(* IEC 61131-3 sources: CS_4_Aufzugsteuerung/src/Stations/CP112/Steuerung/Class/SafetyBaseFSoE (part 6) *)

END_FUNCTION

FUNCTION SafetyBaseFSoE::AddToCache
  VAR_INPUT
    p_SDORequestBuffer 	: ^SDORequReadConfig;
    p_SDOResponseBuffer 	: ^SDORespReadConfig;
  END_VAR

  if p_SDORequestBuffer^.us_Length then
    CachedAddr := p_SDORequestBuffer^.ud_Address;
    CachedSize := p_SDORequestBuffer^.us_Length;
    _memcpy(ptr1:=#Cache, ptr2:=#p_SDOResponseBuffer^.ud_Data, cntr:=p_SDORequestBuffer^.us_Length);
  end_if;

END_FUNCTION

FUNCTION SafetyBaseFSoE::GetFSoEConnectionInfos
  VAR_INPUT
    p_SDORequestBuffer 	: ^SafetyBaseFSoE::SDORequReadConfig;
    p_SDOResponseBuffer 	: ^SafetyBaseFSoE::SDORespReadConfig;
  END_VAR
  VAR
    Address         : UDINT;
    Size            : USINT;
    sd_retval       : DINT;
    i               : UDINT;
    pActConnection  : ^t_FSoEConnectionDetails;
    TempRoutingInfo : t_FSoERoutingInfoElement;
    NextAddress     : UDINT;
  END_VAR

  // always free the connection infos
  FreeFSoEConnectionInfos(bFreeAlways:=TRUE);

  // check if we already got the info:
  if ConnectionInfos.ConnectionNo | ConnectionInfos.pFirstConnection then
    LogError("@0280 (SafetyBaseFSoE::GetFSoEConnectionInfos) List already exists! May not have been resetted correctly!");
    return;
  end_if;

//*****************************************************************************
//** CONNECTION STATE INFO                                                   **
//*****************************************************************************

  // get number of connections
  Address := SBF_SDO_ADDRESS_FSOE_CONN_STATE;
  Size    := 2;

  //send request and receive data
  sd_retval := SDOReadCfgRequ ( p_SDORequestBuffer  := p_SDORequestBuffer
                              , p_SDOResponseBuffer := p_SDOResponseBuffer
                              , ud_Address          := Address
                              , us_Length           := Size
                              );

  //no response
  if ( sd_retval <> 0 ) then
    LogError("@0281 (SafetyBaseFSoE::GetFSoEConnectionInfos) Error reading number of connections.");
    return;
  end_if;

  ConnectionInfos.ConnectionNo := p_SDOResponseBuffer^.ud_Data$UINT;

  if ConnectionInfos.ConnectionNo = 0 then
    // no connections available
    return;
  end_if;

  // allocate memory for the connections
  ConnectionInfos.pFirstConnection$pVoid := ToStdLib.Malloc(size:= ConnectionInfos.ConnectionNo * sizeof(t_FSoEConnectionDetails));

  if ConnectionInfos.pFirstConnection = NIL then
    LogError("@0282 (SafetyBaseFSoE::GetFSoEConnectionInfos) Failed to allocate memory for FSoE connection details.");
    return;
  end_if;

  // reset memory (also resets pNext although we are not using a linked list here)
  _memset(dest:=ConnectionInfos.pFirstConnection, usByte:=0, cntr:= ConnectionInfos.ConnectionNo * sizeof(t_FSoEConnectionDetails));

  Address += Size;
  Size    := 1;

  pActConnection := ConnectionInfos.pFirstConnection;

  // get connection states
  for i := 0 to ConnectionInfos.ConnectionNo-1 do
    // get state of connection

    //send request and receive data
    sd_retval := SDOReadCfgRequ ( p_SDORequestBuffer  := p_SDORequestBuffer
                                , p_SDOResponseBuffer := p_SDOResponseBuffer
                                , ud_Address          := Address
                                , us_Length           := Size
                                );

    //no response
    if ( sd_retval <> 0 ) then
      LogError("@0283 (SafetyBaseFSoE::GetFSoEConnectionInfos) Error reading connection state.");
      return;
    end_if;

    // get connection state
    pActConnection^.ConnectionState := (p_SDOResponseBuffer^.ud_Data$USINT AND 2#0111)$t_FSoEConnectionState;

    // get info if the module is master or slave at this connection
    pActConnection^.Flags.IsMaster  := (p_SDOResponseBuffer^.ud_Data$USINT AND 2#1000) <> 0;

    // save safety number
    pActConnection^.OwnerSafetyNbr  := SafetyNumber;

    // for easier debugging we set the correct next pointers
    if i = ConnectionInfos.ConnectionNo-1 then
      pActConnection^.pNext := NIL;
    else
      pActConnection^.pNext := pActConnection + sizeof(t_FSoEConnectionDetails);
    end_if;

    pActConnection                  += sizeof(t_FSoEConnectionDetails);
    Address                         += Size;
  end_for;

//*****************************************************************************
//** ROUTING INFO                                                            **
//*****************************************************************************

  // get number of connections
  Address := SBF_SDO_ADDRESS_FSOE_ROUTING_INFO;
  Size    := 2;

  //send request and receive data
  sd_retval := SDOReadCfgRequ ( p_SDORequestBuffer  := p_SDORequestBuffer
                              , p_SDOResponseBuffer := p_SDOResponseBuffer
                              , ud_Address          := Address
                              , us_Length           := Size
                              );

  //no response
  if ( sd_retval <> 0 ) then
    LogError("@0281 (SafetyBaseFSoE::GetFSoEConnectionInfos) Error reading number of connections.");
    return;
  end_if;

  // check if it's the same number
  if ConnectionInfos.ConnectionNo <> p_SDOResponseBuffer^.ud_Data$UINT then
    LogError("@0285 (SafetyBaseFSoE::GetFSoEConnectionInfos) Number of connections does not match (case 1).");
    return;
  end_if;

  Address += Size;
  Size    := sizeof(t_FSoERoutingInfoElement);

  pActConnection := ConnectionInfos.pFirstConnection;

  // get connection states
  for i := 0 to ConnectionInfos.ConnectionNo-1 do
    // get routing info of connections

    //send request and receive data
    sd_retval := SDOReadCfgRequ ( p_SDORequestBuffer  := p_SDORequestBuffer
                                , p_SDOResponseBuffer := p_SDOResponseBuffer
                                , ud_Address          := Address
                                , us_Length           := Size
                                );

    //no response
    if ( sd_retval <> 0 ) then
      LogError("@0286 (SafetyBaseFSoE::GetFSoEConnectionInfos) Error reading routing info.");
      return;
    end_if;

    TempRoutingInfo := p_SDOResponseBuffer^.ud_Data$t_FSoERoutingInfoElement;

    // store the data in the connection info
    pActConnection^.SlaveAddress        := TempRoutingInfo.SlaveAddress;
    pActConnection^.MasterReadSize      := TempRoutingInfo.SafeOutputFrameSize;
    pActConnection^.MasterWriteSize     := TempRoutingInfo.SafeInputFrameSize;

    // the offset info depends on if we are master or slave
    if pActConnection^.Flags.IsMaster then
      pActConnection^.MasterReadOffset  := TempRoutingInfo.SafeOutputFrameOffset;
      pActConnection^.MasterWriteOffset := TempRoutingInfo.SafeInputFrameOffset;
    else
      pActConnection^.SlaveWriteOffset  := TempRoutingInfo.SafeOutputFrameOffset;
      pActConnection^.SlaveReadOffset   := TempRoutingInfo.SafeInputFrameOffset;
    end_if;

    pActConnection                  += sizeof(t_FSoEConnectionDetails);
    Address                         += Size;
  end_for;

//*****************************************************************************
//** CONNECTION INSTANCES                                                    **
//*****************************************************************************

  Address := SBF_SDO_ADDRESS_FSOE_CONN_INST;
  Size    := 4;

  //send request and receive data
  sd_retval := SDOReadCfgRequ ( p_SDORequestBuffer  := p_SDORequestBuffer
                              , p_SDOResponseBuffer := p_SDOResponseBuffer
                              , ud_Address          := Address
                              , us_Length           := Size
                              );

  //no response
  if ( sd_retval <> 0 ) then
    LogError("@0281 (SafetyBaseFSoE::GetFSoEConnectionInfos) Error reading number of connections.");
    return;
  end_if;

  // check if it's the same number
  if ConnectionInfos.ConnectionNo <> p_SDOResponseBuffer^.ud_Data then
    LogError("@0287 (SafetyBaseFSoE::GetFSoEConnectionInfos) Number of connections does not match (case 2).");
    return;
  end_if;

  Address += Size;

  pActConnection := ConnectionInfos.pFirstConnection;

  // get connection states
  for i := 0 to ConnectionInfos.ConnectionNo-1 do
    // get routing instance info of connections

    Size := 4;

    //send request and receive data
    sd_retval := SDOReadCfgRequ ( p_SDORequestBuffer  := p_SDORequestBuffer
                                , p_SDOResponseBuffer := p_SDOResponseBuffer
                                , ud_Address          := Address
                                , us_Length           := Size
                                );

    //no response
    if ( sd_retval <> 0 ) then
      LogError("@0288 (SafetyBaseFSoE::GetFSoEConnectionInfos) Error reading size of routing instance info.");
      return;
    end_if;

    // calculate address of next connection (to check it later)
    NextAddress := Address + p_SDOResponseBuffer^.ud_Data;

    // get the flags
    Address   += Size;
    Size      := 4;

    //send request and receive data
    sd_retval := SDOReadCfgRequ ( p_SDORequestBuffer  := p_SDORequestBuffer
                                , p_SDOResponseBuffer := p_SDOResponseBuffer
                                , ud_Address          := Address
                                , us_Length           := Size
                                );

    //no response
    if ( sd_retval <> 0 ) then
      LogError("@0289 (SafetyBaseFSoE::GetFSoEConnectionInfos) Error reading flags of routing instance info.");
      return;
    end_if;

    if ((p_SDOResponseBuffer^.ud_Data AND 1) <> 0) <> pActConnection^.Flags.IsMaster then
      LogError("@028A (SafetyBaseFSoE::GetFSoEConnectionInfos) Master settings mismatch.");
      return;
    end_if;

    //! Flags
    //  Actually, type is 4 bytes in size but for compatibility reasons it is still used as 1 byte. As a result, bits 9-32 are currently not used.
    //  Bit1: 1, wenn FSoE-Master, 0=FSoE-Slave
    //  Bit2: 1, wenn die Slave-Adresse über den HW-Pfad ermittelt wird
    //  Bit3: 1, wenn CRC von der FW ermittelt werden muss
    //  Bit4: 1, wenn Interface und Slave
    //  Bit5: 1, wenn Multichannel verwendet werden, aber ein Multichannel ist nicht vorhanden und der Eingang auf 1 gesetzt wird.
    //  Bit6: 1, wenn der Adressvergabeservice verwendet werden soll
    //  Bit7: 1, wenn der Master beim Slave die Connection ID anfordert
    //  Bit8: 1, wenn es sich um ein HGW handelt
    //  Bit9: 1, wenn Assign Slave On Demand
    //  Bits 10-32: reserviert, sind auf 0 gesetzt und werden nicht ausgewertet

    //check size of FSoEFlags type --> possible are 1 or 4 byte
    pActConnection^.Flags := p_SDOResponseBuffer^.ud_Data$t_FSoEFlags;

    if (pActConnection^.Flags AND SM_FLAGS_FLEXCON_MASK) = SM_FLAGS_FLEXCON_NODE then
#ifdef SAFETY_DEBUG_LOGGING_ACTIVATED
      LogError(e_msg:="SafetyBaseFSoE: Found FSOE Connection of FlexConNode");
#endif
      sFlexCon.FoundNodeInConfig := TRUE;
    elsif (pActConnection^.Flags AND SM_FLAGS_FLEXCON_MASK) = SM_FLAGS_FLEXCON_HOST then
#ifdef SAFETY_DEBUG_LOGGING_ACTIVATED
      LogError(e_msg:="SafetyBaseFSoE: Found FSOE Connection of FlexConHost");
#endif
      sFlexCon.FoundHostInConfig := TRUE;
    end_if;

    // get the net size of the safe output data (only the bits for the I/Os without crc and stuff)
    Address   += Size;
    Size      := 2;

    //send request and receive data
    sd_retval := SDOReadCfgRequ ( p_SDORequestBuffer  := p_SDORequestBuffer
                                , p_SDOResponseBuffer := p_SDOResponseBuffer
                                , ud_Address          := Address
                                , us_Length           := Size
                                );

    //no response
    if ( sd_retval <> 0 ) then
      LogError("@028B (SafetyBaseFSoE::GetFSoEConnectionInfos) Error reading safe output net size of routing instance info.");
      return;
    end_if;

    // we don't need the net size yet

    // get the net size of the safe input data (only the bits for the I/Os without crc and stuff)
    Address   += Size;
    Size      := 2;

    //send request and receive data
    sd_retval := SDOReadCfgRequ ( p_SDORequestBuffer  := p_SDORequestBuffer
                                , p_SDOResponseBuffer := p_SDOResponseBuffer
                                , ud_Address          := Address
                                , us_Length           := Size
                                );

    //no response
    if ( sd_retval <> 0 ) then
      LogError("@028C (SafetyBaseFSoE::GetFSoEConnectionInfos) Error reading safe input net size of routing instance info.");
      return;
    end_if;

    // we don't need the net size yet

    // get the slave address
    Address   += Size;
    Size      := 2;

    //send request and receive data
    sd_retval := SDOReadCfgRequ ( p_SDORequestBuffer  := p_SDORequestBuffer
                                , p_SDOResponseBuffer := p_SDOResponseBuffer
                                , ud_Address          := Address
                                , us_Length           := Size
                                );

    //no response
    if ( sd_retval <> 0 ) then
      LogError("@028D (SafetyBaseFSoE::GetFSoEConnectionInfos) Error reading slave address of routing instance info.");
      return;
    end_if;

    // the following settings are only available in the master
    if pActConnection^.Flags.IsMaster then

      // get the connection ID
      Address   += Size;
      Size      := 2;

      //send request and receive data
      sd_retval := SDOReadCfgRequ ( p_SDORequestBuffer  := p_SDORequestBuffer
                                  , p_SDOResponseBuffer := p_SDOResponseBuffer
                                  , ud_Address          := Address
                                  , us_Length           := Size
                                  );

      //no response
      if ( sd_retval <> 0 ) then
        LogError("@028E (SafetyBaseFSoE::GetFSoEConnectionInfos) Error reading the connection ID of routing instance info.");
        return;
      end_if;

      pActConnection^.ConnectionID := p_SDOResponseBuffer^.ud_Data$UINT;

      // get transmission time
      Address   += Size;
      Size      := 2;

      //send request and receive data
      sd_retval := SDOReadCfgRequ ( p_SDORequestBuffer  := p_SDORequestBuffer
                                  , p_SDOResponseBuffer := p_SDOResponseBuffer
                                  , ud_Address          := Address
                                  , us_Length           := Size
                                  );

      //no response
      if ( sd_retval <> 0 ) then
        LogError("@028F (SafetyBaseFSoE::GetFSoEConnectionInfos) Error reading the transmission time of routing instance info.");
        return;
      end_if;

      pActConnection^.TransmissionTime_ms := p_SDOResponseBuffer^.ud_Data$UINT;

      // get length of communication parameters (must be 2)
      Address   += Size;
      Size      := 2;

      //send request and receive data
      sd_retval := SDOReadCfgRequ ( p_SDORequestBuffer  := p_SDORequestBuffer
                                  , p_SDOResponseBuffer := p_SDOResponseBuffer
                                  , ud_Address          := Address
                                  , us_Length           := Size
                                  );

      //no response
      if ( sd_retval <> 0 ) then
        LogError("@0290 (SafetyBaseFSoE::GetFSoEConnectionInfos) Error reading the length of the communication parameters of routing instance info.");
        return;
      end_if;

      if p_SDOResponseBuffer^.ud_Data$UINT <> 2 then
        LogError("@0291 (SafetyBaseFSoE::GetFSoEConnectionInfos) Length of communication parameters is wrong.");
        return;
      end_if;

      // skip FSoE watchdog time in ms
      Address   += Size;
      Size      := 2;

      // get size of application parameters
      Address   += Size;
      Size      := 2;

      //send request and receive data
      sd_retval := SDOReadCfgRequ ( p_SDORequestBuffer  := p_SDORequestBuffer
                                  , p_SDOResponseBuffer := p_SDOResponseBuffer
                                  , ud_Address          := Address
                                  , us_Length           := Size
                                  );

      //no response
      if ( sd_retval <> 0 ) then
        LogError("@0292 (SafetyBaseFSoE::GetFSoEConnectionInfos) Error reading the length of the application parameters of routing instance info.");
        return;
      end_if;

      // skip length
      Address   += Size;

      // skip application parameters
      Size      := p_SDOResponseBuffer^.ud_Data$USINT;
      Address   += Size;

      // get to a 4 byte aligned address
      if (Address MOD 4) then
        Address := Address + (4 - (Address MOD 4)); //increase memory, up to a value, which could be divided by 4
      end_if;

      // get size of hw path
      Size      := 4;

      //send request and receive data
      sd_retval := SDOReadCfgRequ ( p_SDORequestBuffer  := p_SDORequestBuffer
                                  , p_SDOResponseBuffer := p_SDOResponseBuffer
                                  , ud_Address          := Address
                                  , us_Length           := Size
                                  );

      //no response
      if ( sd_retval <> 0 ) then
        LogError("@0293 (SafetyBaseFSoE::GetFSoEConnectionInfos) Error reading the hardware path length of routing instance info.");
        return;
      end_if;

      // get the hardware path
      Address   += Size;
      Size      := p_SDOResponseBuffer^.ud_Data$USINT;

      if Size = 0 then
        LogError("@0294 (SafetyBaseFSoE::GetFSoEConnectionInfos) Hardware path length is zero.");
        return;
      end_if;

      //send request and receive data
      sd_retval := SDOReadCfgRequ ( p_SDORequestBuffer  := p_SDORequestBuffer
                                  , p_SDOResponseBuffer := p_SDOResponseBuffer
                                  , ud_Address          := Address
                                  , us_Length           := Size
                                  );

      //no response
      if ( sd_retval <> 0 ) then
        LogError("@0295 (SafetyBaseFSoE::GetFSoEConnectionInfos) Error reading the hardware path of routing instance info.");
        return;
      end_if;

      // save hardware path into structure
      pActConnection^.SlavePathLen      := Size;
      pActConnection^.pSlavePath$pVoid  := ToStdLib.Malloc(size:=Size);

      if pActConnection^.pSlavePath = NIL then
        LogError("@0296 (SafetyBaseFSoE::GetFSoEConnectionInfos) Failed to allocate memory for the slave hardware path at the routing instance info.");
        return;
      end_if;

      _memcpy(ptr1:=pActConnection^.pSlavePath, ptr2:=#p_SDOResponseBuffer^.ud_Data, cntr:=pActConnection^.SlavePathLen);

      Address         += Size;

      // get to a 4 byte aligned address
      if (Address MOD 4) then
        Address := Address + (4 - (Address MOD 4)); //increase memory, up to a value, which could be divided by 4
      end_if;

      // get size of compressed hw path
      Size      := 4;

      //send request and receive data
      sd_retval := SDOReadCfgRequ ( p_SDORequestBuffer  := p_SDORequestBuffer
                                  , p_SDOResponseBuffer := p_SDOResponseBuffer
                                  , ud_Address          := Address
                                  , us_Length           := Size
                                  );

      //no response
      if ( sd_retval <> 0 ) then
        LogError("@0297 (SafetyBaseFSoE::GetFSoEConnectionInfos) Error reading the compressed hardware path length of routing instance info.");
        return;
      end_if;

      // get the hardware path
      Address   += Size;
      Size      := p_SDOResponseBuffer^.ud_Data$USINT;

      //send request and receive data
      sd_retval := SDOReadCfgRequ ( p_SDORequestBuffer  := p_SDORequestBuffer
                                  , p_SDOResponseBuffer := p_SDOResponseBuffer
                                  , ud_Address          := Address
                                  , us_Length           := Size
                                  );

      //no response
      if ( sd_retval <> 0 ) then
        LogError("@0298 (SafetyBaseFSoE::GetFSoEConnectionInfos) Error reading the compressed hardware path of routing instance info.");
        return;
      end_if;

      // save compressed hardware path into structure
      pActConnection^.SlavePathCompLen      := Size;
      pActConnection^.pSlavePathComp$pVoid  := ToStdLib.Malloc(size:=Size);

      if pActConnection^.pSlavePathComp = NIL then
        LogError("@0299 (SafetyBaseFSoE::GetFSoEConnectionInfos) Failed to allocate memory for the compressed slave hardware path at the routing instance info.");
        return;
      end_if;

      _memcpy(ptr1:=pActConnection^.pSlavePathComp, ptr2:=#p_SDOResponseBuffer^.ud_Data, cntr:=pActConnection^.SlavePathCompLen);

      if  (pActConnection^.pSlavePathComp^ = 6) &
          ((pActConnection^.pSlavePathComp + 5)^$HDINT AND 16#00FFFFFF) = 0 then

        // special IP: (0.0.0.x)
        // if custom ip is detected change pathcomp type from 6 (IP) to 3 (Interface)
        pActConnection^.pSlavePathComp^ :=3;
      end_if;

      //Get slot ID and communication ID from HGW
      if pActConnection^.Flags.IsHGW then

        //Get machinenumber of FUB
        sd_retval := SDOReadCfgRequ ( p_SDORequestBuffer  := p_SDORequestBuffer
                                    , p_SDOResponseBuffer := p_SDOResponseBuffer
                                    , ud_Address          := SBF_SDO_ADDRESS_HGW_FUB_BASE_ADDRESS + SBF_SDO_ADDRESS_HGW_OFFSET_MACHINENUMBER
                                    , us_Length           := 4
                                    , b_UseCache          := FALSE
                                    );

        //no response
        if ( sd_retval <> 0 ) then
          LogError("@03DA (SafetyBaseFSoE::GetFSoEConnectionInfos) Error reading the machinenumber of routing instance info.");
          return;
        end_if;

        sHGW.udMachineNrb := p_SDOResponseBuffer^.ud_Data$UDINT;

        // get the Slot ID
        Address   += Size;
        Size      := 2;

        //send request and receive data
        sd_retval := SDOReadCfgRequ ( p_SDORequestBuffer  := p_SDORequestBuffer
                                    , p_SDOResponseBuffer := p_SDOResponseBuffer
                                    , ud_Address          := Address
                                    , us_Length           := Size
                                    );

        //no response
        if ( sd_retval <> 0 ) then
          LogError("@03DB (SafetyBaseFSoE::GetFSoEConnectionInfos) Error reading the communication ID of routing instance info.");
          return;
        end_if;

        sHGW.uiCommunicationID := p_SDOResponseBuffer^.ud_Data$UINT;

        // get the communication ID
        Address   += Size;
        Size      := 2;

        //send request and receive data
        sd_retval := SDOReadCfgRequ ( p_SDORequestBuffer  := p_SDORequestBuffer
                                    , p_SDOResponseBuffer := p_SDOResponseBuffer
                                    , ud_Address          := Address
                                    , us_Length           := Size
                                    );

        //no response
        if ( sd_retval <> 0 ) then
          LogError("@03DC (SafetyBaseFSoE::GetFSoEConnectionInfos) Error reading the slot ID of routing instance info.");
          return;
        end_if;

        sHGW.uiSlotID := p_SDOResponseBuffer^.ud_Data$UINT;

        //save fsoe pdo offsets and length
        sHGW.InputPDOLength  := pActConnection^.MasterWriteSize;
        sHGW.OutputPDOLength := pActConnection^.MasterReadSize;
        if pActConnection^.Flags.IsMaster then
          sHGW.InputPDOOffset  := pActConnection^.MasterWriteOffset;
          sHGW.OutputPDOOffset := pActConnection^.MasterReadOffset;
        else
          sHGW.InputPDOOffset  := pActConnection^.SlaveWriteOffset;
          sHGW.OutputPDOOffset := pActConnection^.SlaveReadOffset;
        end_if;
        sHGW.uiTransmissionTime_ms := pActConnection^.TransmissionTime_ms;
      end_if;

      Address         += Size;

      // get to a 4 byte aligned address
      if (Address MOD 4) then
        Address := Address + (4 - (Address MOD 4)); //increase memory, up to a value, which could be divided by 4
      end_if;

      if Address > NextAddress then
        LogError("@029A (SafetyBaseFSoE::GetFSoEConnectionInfos) Structure size mismatch.");
        return;
      end_if;
    end_if;

    Address         := NextAddress;
    pActConnection  += sizeof(t_FSoEConnectionDetails);
  end_for;

END_FUNCTION

FUNCTION SafetyBaseFSoE::FreeFSoEConnectionInfos
	VAR_INPUT
		bFreeAlways 	: BOOL;(* := false *)
	END_VAR
  VAR
    i               : UDINT;
    pActConnection  : ^t_FSoEConnectionDetails;
  END_VAR

  if (ConnectionInfos.ConnectionNo = 0) | (ConnectionInfos.pFirstConnection = NIL) then
    // nothing to free
    return;
  end_if;

  //Check if we want to clear the connection infos always
  if bFreeAlways = false then
    // check if all connections have been initialized
    pActConnection := ConnectionInfos.pFirstConnection;
    for i := 0 to ConnectionInfos.ConnectionNo-1 do
      if pActConnection^.ConnectionState = FCS_NOT_INITIALIZED then
        // not yet time to free them
        return;
      end_if;

      pActConnection += sizeof(t_FSoEConnectionDetails);
    end_for;
  end_if;

  pActConnection := ConnectionInfos.pFirstConnection;
  for i := 0 to ConnectionInfos.ConnectionNo-1 do
    // free hardware path memory

    if pActConnection^.pSlavePath then
      ToStdLib.Free(mptr:=pActConnection^.pSlavePath);
    end_if;

    if pActConnection^.pSlavePathComp then
      ToStdLib.Free(mptr:=pActConnection^.pSlavePathComp);
    end_if;

    pActConnection += sizeof(t_FSoEConnectionDetails);
  end_for;

  // free the connectionlist
  ToStdLib.Free(mptr:=ConnectionInfos.pFirstConnection);
  ConnectionInfos.pFirstConnection := NIL;
  ConnectionInfos.ConnectionNo := 0;

END_FUNCTION

FUNCTION SafetyBaseFSoE::CheckFSoEConnections
  VAR
    MyPara 	            : CmdStruct;
    MyResult	          : results;
    i                   : UDINT;
    pActConnection      : ^t_FSoEConnectionDetails;
    SDORequestBuffer    : SDORequReadConfig;
    SDOResponseBuffer   : ARRAY [0..SBF_SDO_MAX_LENGTH-1] OF USINT;
    p_SDORequestBuffer 	: ^SDORequReadConfig;
    p_SDOResponseBuffer : ^SDORespReadConfig;
    UnInifializedNo     : UDINT;
    sd_retval           : DINT;
  END_VAR

  // there were some of the FSoE connections not initialized when fetching the configuration data => update them

  UnInifializedNo := 0;

  //SDO request for this command has 5 bytes additional to the header
  p_SDORequestBuffer := #SDORequestBuffer;

  //SDO response for this command can have maximum additional data
  p_SDOResponseBuffer := (#SDOResponseBuffer)$^SDORespReadConfig;

  //calculate length without crc
  p_SDORequestBuffer^.StdHeader.Len := sizeof(SDORequReadConfig) - sizeof(SDOHeader.StdHeader.CRC);

  //type
  p_SDORequestBuffer^.StdHeader.Typ := SDO_STD;

  //command for reading config data
  p_SDORequestBuffer^.StdHeader.Cmd := SBF_SDO_COMMAND_READ;

  // reset cache, because it may contain an old access on the same address => we want fresh data
  CachedSize := 0;

  pActConnection := ConnectionInfos.pFirstConnection;

  for i := 0 to ConnectionInfos.ConnectionNo-1 do
    if pActConnection^.ConnectionState = FCS_NOT_INITIALIZED then
      UnInifializedNo += 1;

      //send request and receive data
      sd_retval := SDOReadCfgRequ ( p_SDORequestBuffer  := p_SDORequestBuffer
                                  , p_SDOResponseBuffer := p_SDOResponseBuffer
                                  , ud_Address          := SBF_SDO_ADDRESS_FSOE_CONN_STATE + 2 + i
                                  , us_Length           := 1
                                  );

      //no response
      if ( sd_retval <> 0 ) then
        LogError("@0283 (SafetyBaseFSoE::CheckFSoEConnections) Error reading connection state.");
        return;
      end_if;

      // get connection state
      pActConnection^.ConnectionState := (p_SDOResponseBuffer^.ud_Data$USINT AND 2#0111)$t_FSoEConnectionState;

      if pActConnection^.ConnectionState <> FCS_NOT_INITIALIZED then
        UnInifializedNo -= 1;

        // get the corresponding slave address number

        //send request and receive data
        sd_retval := SDOReadCfgRequ ( p_SDORequestBuffer  := p_SDORequestBuffer
                                    , p_SDOResponseBuffer := p_SDOResponseBuffer
                                    , ud_Address          := SBF_SDO_ADDRESS_FSOE_ROUTING_INFO + 2 + i * sizeof(t_FSoERoutingInfoElement)
                                    , us_Length           := sizeof(t_FSoERoutingInfoElement)
                                    );

        //no response
        if ( sd_retval <> 0 ) then
          LogError("@0286 (SafetyBaseFSoE::CheckFSoEConnections) Error reading routing info.");
          return;
        end_if;

        pActConnection^.SlaveAddress := p_SDOResponseBuffer^.ud_Data$t_FSoERoutingInfoElement.SlaveAddress;

        if pActConnection^.SlaveAddress = 0 then
          LogError("@029B (SafetyBaseFSoE::CheckFSoEConnections) Connection initialized but slave address is still zero!");
        end_if;
      end_if;
    end_if;

    pActConnection                  += sizeof(t_FSoEConnectionDetails);
  end_for;

  // if all connections are initialized => tell the safety manager
  if (UnInifializedNo = 0) & pSafetyManagerThis then
    MyPara.uiCmd    := CMD_SM_FSOE_CON_INITIALIZED;
    MyPara.aPara[0] := SafetyNumber$DINT;
    MyPara.aPara[1] := ConnectionInfos.ConnectionNo$DINT;
    MyPara.aPara[2] := ConnectionInfos.pFirstConnection$DINT;

    if pSafetyManagerThis^.NewInst(#MyPara, #MyResult) = READY then
      // we don't need this memory anymore
      FreeFSoEConnectionInfos();
    end_if;
  end_if;

END_FUNCTION

FUNCTION VIRTUAL GLOBAL SafetyBaseFSoE::GetDiagConnect::NewInst
  VAR_INPUT
    pPara 	: ^CmdStruct;
    pResult 	: ^Results;
  END_VAR
  VAR_OUTPUT
    ret_code 	: IprStates;
  END_VAR

  ret_code := READY;

  CASE pPara^.uiCmd OF

    CMD_SM_DIAG_GET_INFO:

      //Subcommand
      case pPara^.aPara[0] of
//*****************************************************************************
        SBCMD_SM_DIAG_GET_INFO:
          pResult^.aData[0] :=  GetDiagInfo(pDiagInfo:=(pPara^.aPara[1])$^SafetyDiagInfo);

//*****************************************************************************
        SBCMD_SM_DIAG_GET_STATE:
          pResult^.aData[0] :=  GetDiagState(pDiagState:=(pPara^.aPara[1])$^SafetyDiagState);

//*****************************************************************************
        SBCMD_SM_DIAG_FETCH_INFO:
      //Fetch Diag Info for uCx
          FetchDiagInfo(ucChoice:=pPara^.aPara[1]$USINT);

//*****************************************************************************
        SBCMD_SM_DIAG_FETCH_STATE:
          FetchDiagState();

//*****************************************************************************
        SBCMD_SM_DIAG_IS_SAVE_LOG_ACTIVE:
          pResult^.aData[0] := SaveLogActive();

//*****************************************************************************
        SBCMD_SM_DIAG_SAVE_LOGFILE:
          pResult^.aData[0] := (SaveLog(ucChoice:=(pPara^.aPara[1])$USINT, pDPNE:=(pPara^.aPara[2])$^CHAR))$USINT;

//*****************************************************************************
        SBCMD_SM_DIAG_GET_SAVE_LOGFILE_STATE:
          pResult^.aData[0] := DiagVars.SavingLogSuccessful$USINT;

//*****************************************************************************
        SBCMD_SM_DIAG_GET_SAFETY_NUMBER:
          pResult^.aData[0]$UDINT := SafetyNumber;

//*****************************************************************************
        SBCMD_SM_DIAG_GET_SAFETY_STATE:
          pResult^.aData[0] := SafetyState$USINT;

//*****************************************************************************
        SBCMD_SM_DIAG_IS_DIAGNOSE_AVAILABLE:
          pResult^.aData[0] := TRUE;

//*****************************************************************************
        SBCMD_SM_DIAG_GET_CHANNEL_INFO:
          pResult^.aData[0] := GetChannelInfo(pErrorMemUser:=(pPara^.aPara[1])$^UINT, pErrorMem:=#aErrorMem[1], ErrorDataLength:=aErrorMem[0] - 1);
          pResult^.aData[1] := aErrorMem[0] - 1;

//*****************************************************************************
        SBCMD_SM_DIAG_FETCH_CHANNEL_INFO:
          FetchChannelInfo();

//*****************************************************************************
        SBCMD_SM_DIAG_GET_ERRORCODE_OFFSET:

          //Check for valid version
          if pPara^.aPara[1] = 0x01 then  //Version

            ret_code := READY;
            pResult^.aData[0] := 0x01;  //return version
            pResult^.aData[1]$UDINT := GetDiagVisualOffsetErrorCode();

            pResult^.uiLng := 12;

          else

            //invalid version, return error
            ret_code := ERROR;

            pResult^.aData[0] := 0x0;
            pResult^.uiLng    := 4;

          end_if;

        END_CASE;
    else
      TRACE("(SafetyBaseFSoE::GetDiagConnect::NewInst) Unknown command!");
      ret_code := ERROR;
  END_CASE;

END_FUNCTION

FUNCTION SafetyBaseFSoE::GetNewMemSize
  VAR_INPUT
    Required 	: UDINT;
  END_VAR
  VAR_OUTPUT
    NextBiggerBlockSize 	: UDINT;
  END_VAR

  // how many complete blocks are necessary
  NextBiggerBlockSize := Required / SBF_CONFIG_MEMORY_BLOCK_SIZE;

  // is there also an incomplete block?
  if Required MOD SBF_CONFIG_MEMORY_BLOCK_SIZE then
    NextBiggerBlockSize += 1;
  end_if;

  // now that we have the number of blocks necessary => get number of bytes
  NextBiggerBlockSize *= SBF_CONFIG_MEMORY_BLOCK_SIZE;

END_FUNCTION

FUNCTION SafetyBaseFSoE::CheckAddDynSlaveResponse
  VAR_INPUT
    pAddDynSlaveRsp 	: ^t_AddDynSlaveResponse;
  END_VAR
  VAR_OUTPUT
    ResponseOk 	: BOOL;
  END_VAR

  // check if any of the offset/length combination exceeds our access to the module
  if ((pAddDynSlaveRsp^.OffsetSafeInData  + pAddDynSlaveRsp^.LenSafeInData ) > MyPDOWriteSize) |
     ((pAddDynSlaveRsp^.OffsetSafeOutData + pAddDynSlaveRsp^.LenSafeOutData) > MyPDOReadSize ) then
    ResponseOk := FALSE;

    LogError("@029C (SafetyBaseFSoE::CheckAddDynSlaveResponse) Invalid offset/length combination of read or write data in AddDynSlave response.");
  else
    ResponseOk := TRUE;
  end_if;

END_FUNCTION

FUNCTION SafetyBaseFSoE::GetChannelInfo
  VAR_INPUT
    pErrorMemUser 	: ^UINT;
    pErrorMem 	: ^USINT;
    ErrorDataLength 	: INT;
  END_VAR
  VAR_OUTPUT
    StateReady 	: BOOL;
  END_VAR
  VAR
    i   : INT;
  END_VAR

  StateReady := DiagVars.UserErrorInfoReady;

  if StateReady then
    //copy error values in UserArray
    for i := 0 to ErrorDataLength-1 do

      pErrorMemUser^ := pErrorMem^;

      if (pErrorMemUser^ <> 0) then
        pErrorMemUser^ += GetDiagVisualOffsetErrorCode()$UINT; //Add offset to each errorvalue so that it matches the value in SafetyDesigner.
      end_if;

      //set pointer to next entry
      pErrorMemUser += sizeof(UINT);
      pErrorMem += sizeof(USINT);
    end_for;
  end_if;

END_FUNCTION

FUNCTION VIRTUAL GLOBAL SafetyBaseFSoE::FetchChannelInfo

  DiagVars.UserErrorInfoReady := FALSE;
  DiagVars.UserWantsErrorInfo := TRUE;

END_FUNCTION

#pragma warning(disable:73);
FUNCTION VIRTUAL SafetyBaseFSoE::SafeActModuleConfig
  VAR_INPUT
    sActModuleConfig 	: t_ModuleCfg;
  END_VAR
  //overwrite this function at derived class to safe module config
END_FUNCTION
#pragma warning(default:73);

FUNCTION VIRTUAL SafetyBaseFSoE::GetDiagVisualOffsetErrorCode
	VAR_OUTPUT
		udOffset 	: UDINT;
	END_VAR

  //In the safety firmware for the CSCP and SCP there is only one byte for the errorcode
  //To have different errorcodes (between CSCP and SCP) the safetydesigner adds a fix offset of 1000 to the errorcodes of the SCP01x and SCP11x
  udOffset := 1000;

END_FUNCTION

FUNCTION VIRTUAL SafetyBaseFSoE::AddFastUnsafeRoutElement
	VAR_INPUT
		pRoutTable 	: ^pUnsafeIORoutingElement;
		pRoutElementsNo 	: ^UINT;
		ud_Address 	: UDINT;
		ui_NameLen 	: UINT;
		pNameNewElement 	: ^CHAR;
		BitMask 	: BDINT;(* := 0 *)
		bWriteVar 	: BOOL;
	END_VAR
	VAR_OUTPUT
		sd_retval 	: DINT;
	END_VAR
  VAR
    p_RoutElement   : ^UnsafeIORoutingElement;
  END_VAR

  sd_retval := -1;

  // check parameters
  if (ui_NameLen = 0) | (pNameNewElement = NIL) then
    LogError("@0240 (SafetyBaseFSoE::AddFastUnsafeRoutElement) Invalid call parameters for the variable name (invalid configuration in safety cpu).");
    return;
  end_if;

  //With the first element, the table must be positioned
  if ( pRoutTable^ = NIL ) then

    //allocate memory for first routing element
    pRoutTable^$^void := ToStdLib.Malloc(size := sizeof(UnsafeIORoutingElement));

    if ( pRoutTable^ = NIL ) then

      sd_retval                         := -1;
      SetSafetyState(NewState:=_MemAllocFailed);
      return;

    end_if;

    p_RoutElement := pRoutTable^;

  else

    //add new element

    pRoutTable^$^void := ToStdLib.ReAlloc(mptr := pRoutTable^, newsize := ( ( pRoutElementsNo^ + 1 ) * sizeof(UnsafeIORoutingElement)));

    if ( pRoutTable^ = NIL ) then

      sd_retval                         := -1;
      SetSafetyState(NewState:=_MemAllocFailed);
      return;

    end_if;

    //set pointer to empty element on last position
    p_RoutElement := pRoutTable^ + ( pRoutElementsNo^ ) * sizeof(UnsafeIORoutingElement);

  end_if;

  if p_RoutElement then
    //allocate memory for name
    p_RoutElement^.pName$^void := ToStdLib.Malloc(size := ui_NameLen);

    if ( p_RoutElement^.pName = NIL ) then

      sd_retval                         := -1;
      SetSafetyState(NewState:=_MemAllocFailed);
      return;

    end_if;

    p_RoutElement^.NameLength := ui_NameLen;
    _memcpy(ptr1:=p_RoutElement^.pName, ptr2:=pNameNewElement, cntr:=ui_NameLen);

    p_RoutElement^.BitMask := BitMask;

    // initialize with invalid
    p_RoutElement^.b_IsValid            := FALSE;
    p_RoutElement^.sd_OldValue          := (16#80000000)$DINT;
    p_RoutElement^.sd_NewValue4External := (16#80000000)$DINT;

    // remember that we haven't transmitted this value so far
    p_RoutElement^.b_AlreadyTransmitted := FALSE;

    if (aFastUnsafeReadDOs[0].pData <> NIL) | (aFastUnsafeWriteDOs[0].pData <> NIL) then

      //check if it's a write or read variable
      if bWriteVar = TRUE then
        //add output variable
        if pFastUnsafeOutBuffer then
          p_RoutElement^.ud_Address := pFastUnsafeOutBuffer$UDINT + ud_Address;
        else
          LogError("@0788 (SafetyBaseFSoE::AddFastUnsafeRoutElement) Add Fast output Variable failed. Invalid Outputbuffer.");
          return;
        end_if;

      else
        //add Input variable
        if pFastUnsafeInBuffer then
          p_RoutElement^.ud_Address := pFastUnsafeInBuffer$UDINT + ud_Address;
        else
          LogError("@0789 (SafetyBaseFSoE::AddFastUnsafeRoutElement) Add Fast input Variable failed. Invalid Inputbuffer.");
          return;
        end_if;

      end_if;
    end_if;

    // initialize next pointer
    p_RoutElement^.pNext := NIL;

    // check if name exists in PLC
    p_RoutElement^.ud_Thisp   := GetThisViaServerName(pNameNewElement)$UDINT;
    if (pRoutTable = #p_UnsafeOutputsTable) & p_RoutElement^.BitMask then
      p_RoutElement^.UnsafeType := BDINTOutput;
    else
      p_RoutElement^.UnsafeType := NormalUnsafe;
    end_if;

    //increase counter
    pRoutElementsNo^ += 1;
  end_if;

END_FUNCTION

FUNCTION VIRTUAL SafetyBaseFSoE::UpdateSafetyNbrAtRoutingElement
	VAR_INPUT
		PathLen 	: UINT;
		pCompressedPath 	: ^USINT;
		SafetyNbr 	: HDINT;
	END_VAR
	VAR_OUTPUT
		Retval 	: DINT;
	END_VAR
  VAR
  	pRoutElement : ^RoutElement;
    i                 : UINT;
  END_VAR

  // initialize the retcode with error
  Retval := -1;

  // check if the path is among our routing elements

  //check each element
  if ( ui_CntRoutElements > 0 ) then
    //set pointer on first routing element
    pRoutElement := p_RoutTable;

    for i := 0 to (ui_CntRoutElements - 1) do

      // if there's a path and the length matches
      if pRoutElement^.p_CompressedPath & (pRoutElement^.ui_ComprPathLen = PathLen) then

        // check the path content
        if ToStdLib.MemCmp(dest:=pCompressedPath, source:=pRoutElement^.p_CompressedPath , size:=PathLen) = 0 then

          // if it's the correct path, set the new safety number for that object
          pRoutElement^.ud_SafeNumber := SafetyNbr;

          // success
          Retval := 0;
          return;

        end_if;
      end_if;

      //set pointer to next element
      pRoutElement += sizeof ( RoutElement );
    end_for;
  end_if;

END_FUNCTION

FUNCTION VIRTUAL GLOBAL SafetyBaseFSoE::QuitError
	VAR_INPUT
		Mode 	: DINT;
	END_VAR
	VAR_OUTPUT
		Retval 	: DINT;
	END_VAR

  case Mode of
//**********************************************************************************************************************************************************
    0: // compatibility mode for SCP111 (if quit error via DLL available, use it with submodules. otherwise use the "only quit comm errors" variant)
      if QuitErrorAvailable then
        // initialize the parameter for compatible behavior (quit with submodules)
        QuitErrorParameter := 1;

        // remember to do it in next background
        QuitComError := 2;
      else
        // remember. that there has been a manual quit (for writing PDOs in PostScan)
        b_ManualQuit := TRUE;

        // remember to do it in next cyclic
        QuitComError := 1;
      end_if;

//**********************************************************************************************************************************************************
    1: // only quit the communication errors (send set bus ready signal)

      // remember. that there has been a manual quit (for writing PDOs in PostScan)
      b_ManualQuit := TRUE;

      // remember to do it in next cyclic
      QuitComError := 1;

//**********************************************************************************************************************************************************
    2: // quit error with submodules

      // check if the function is supported by the CIL interface
      if QuitErrorAvailable then
        // initialize the parameter to quit with submodules
        QuitErrorParameter := 1;

        // remember to do it in next background
        QuitComError := 2;
      else
        // function not available
        QuitComError := -8;
      end_if;

//**********************************************************************************************************************************************************
    3: // quit error without submodules (the current module only)

      // check if the function is supported by the CIL interface
      if QuitErrorAvailable then
        // initialize the parameter to quit without submodules
        QuitErrorParameter := 0;

        // remember to do it in next background
        QuitComError := 3;
      else
        // function not available
        QuitComError := -8;
      end_if;

//**********************************************************************************************************************************************************
  else
    // invalid mode selected
    QuitComError := -7;
  end_case;

  // refresh the server on the outer object
  RefreshAsySrv();

  // return the current server value
  Retval := QuitComError;

END_FUNCTION
